Fanuc KAREL source: kx00029.KL

-- PROVISIONAL review KL for V1013-1; original PC SHA256 4fcdaff24ab3127ebcaf4fcb7661847b13b2ef2193959889d008b5f533b6174f
-- Incomplete behavior may be omitted. Consult companion uncertainty JSON. Do not deploy.
PROGRAM KX00029
%NOLOCKGROUP
VAR
  I : INTEGER
  J : INTEGER
  B : BOOLEAN
  F : FILE
  S : STRING[80]
-- UNRESOLVED_DECL P type=000102
BEGIN
  -- UNRESOLVED_PC offsets 5-12; opcodes 9D,23
  -- UNRESOLVED_PC offsets 17-21; opcodes 7F
END KX00029
